(* IEC 61131-3 sources: 2026_Projet_YGO_ExcavatriceDragage/ARCHIVES/Code/PLC_TESTS/TYPES/STRUCTS, 13 files *)

(* ---- ST_PlcTestsCmd.st ---- *)
// ═══════════════════════════════════════════════════════════════
// 🧪 ST_PlcTestsCmd — Commandes de pilotage du banc de validation
// ═══════════════════════════════════════════════════════════════

TYPE ST_PlcTestsCmd :
STRUCT
    // Commandes unitaires : une seule suite manuelle à la fois.
    RunSafety     : BOOL;   // Lance la suite Safety
    RunTranslation: BOOL;   // Lance la suite Translation
    RunBucket     : BOOL;   // Lance la suite Benne
    RunEncoder    : BOOL;   // Lance la suite Codeurs/Homing
    RunModes      : BOOL;   // Lance la suite Modes/Homme-mort
    RunHeartbeat  : BOOL;   // Lance la suite Heartbeat IHM↔PLC
    RunSupervision: BOOL;   // Lance la suite Supervision/Persistance config
    RunFramework  : BOOL;   // Lance l'autotest indépendant du framework
    RunAll        : BOOL;   // Lance Safety→Translation→Bucket→Encoder→Modes→Heartbeat
    RunSuite      : INT;    // Compatibilité : >0 lance une suite manuelle
    RunCase       : INT;    // Cas de la commande unitaire sélectionnée
    Abort         : BOOL;   // Abandonne le test en cours
    ClearReport   : BOOL;   // Efface les rapports de tests
END_STRUCT
END_TYPE

(* ---- ST_PlcTestsStatus.st ---- *)
// ═══════════════════════════════════════════════════════════════
// 🧪 ST_PlcTestsStatus — États et progression des tests
// ═══════════════════════════════════════════════════════════════

TYPE ST_PlcTestsStatus :
STRUCT
    RunState         : E_TestRunState;
    SimulationActive : BOOL;       // TRUE si la simulation automate est active
    ActiveSuiteId    : INT;        // ID de la suite en cours (ex: 1)
    ActiveCaseId     : INT;        // ID du cas en cours
    ActiveStepId     : INT;        // ID de l'étape en cours
    ActiveSuiteName  : STRING(32); // Nom de la suite active
    ActiveCaseName   : STRING(32); // Nom du cas active
    ActiveStepName   : STRING(32); // Nom de l'étape active
    StepElapsed      : TIME;       // Temps écoulé dans l'étape active
    StepTimeoutPT    : TIME;       // Timeout de l'étape active
    CasesTotal       : INT;        // Nombre total de cas à jouer
    CasesPassed      : INT;        // Nombre de cas réussis
    CasesFailed      : INT;        // Nombre de cas en échec
    Heartbeat        : BOOL;       // Clignotant d'activité (3 pulses sur transition)
    FailureSummary   : STRING(255); // 🏷️ Détail des défauts du dernier run, TOUTES suites confondues (remonte Report.FailureSummary de chaque suite exécutée) — lisible sans creuser Suite*Validation
    TerminalState    : E_TestTerminalState;
    ErrorCode        : INT;
    ErrorMessage     : STRING(160);
    SuiteElapsed     : TIME;
    SuiteWatchdogExpired : BOOL;
END_STRUCT
END_TYPE

(* ---- ST_TestCaseConfig.st ---- *)
// ═══════════════════════════════════════════════════════════════
// 🧪 ST_TestCaseConfig — Configuration d'un cas de test
// ═══════════════════════════════════════════════════════════════

TYPE ST_TestCaseConfig :
STRUCT
    Name      : STRING(32);          // Libellé (ex. 'TC-01 Armement nominal')
    FirstStep : INT;                 // Première étape (SETUP) du cas de test
END_STRUCT
END_TYPE

(* ---- ST_TestCaseResult.st ---- *)
// ═══════════════════════════════════════════════════════════════
// 🧪 ST_TestCaseResult — Résultat d'un cas de test
// ═══════════════════════════════════════════════════════════════

TYPE ST_TestCaseResult :
STRUCT
    Name         : STRING(32);       // 🏷️ Libellé lisible (copié de CaseTable[i].Name) — identifie le cas sans chercher l'index
    Executed     : BOOL;             // Le cas de test a-t-elle été exécuté (ex. non exécuté si setup précédent abort)
    Ok           : BOOL;             // Succès global du cas de test
    FailedStepId : INT;              // Index de la première étape en échec (0 si aucune)
    FailReason   : E_TestFailReason; // Cause de l'échec global du cas de test
    Duration     : TIME;             // Durée totale du cas de test
END_STRUCT
END_TYPE

(* ---- ST_TestCheckConfig.st ---- *)
// ═══════════════════════════════════════════════════════════════
// 🧪 ST_TestCheckConfig — Configuration d'un check (une assertion)
// ═══════════════════════════════════════════════════════════════

TYPE ST_TestCheckConfig :
STRUCT
    Kind         : E_TestCheckKind;  // Type de check
    Mode         : E_TestCheckMode;  // Mode d'évaluation
    ProbeIdx     : INT;              // Index de la sonde dans le tableau correspondant
    ExpectedBool : BOOL;             // Valeur attendue pour BOOL_EQUAL
    ExpectedDint : DINT;             // Valeur attendue pour DINT_EQUAL / DINT_NOT_EQUAL
    ExpectedMin  : DINT;             // Bornes pour DINT_IN_RANGE
    ExpectedMax  : DINT;
    Mask         : WORD;             // Masque pour WORD_MASK_*
    RealMin      : REAL;             // Bornes pour REAL_IN_RANGE
    RealMax      : REAL;
    StablePT     : TIME;             // Durée de stabilité requise pour CHECK_WAIT_UNTIL
END_STRUCT
END_TYPE

(* ---- ST_TestEvent.st ---- *)
// 🧪 Événement journalisé par le banc de test
TYPE ST_TestEvent :
STRUCT
    Sequence       : UDINT;
    Severity       : E_TestEventSeverity;
    SuiteId        : INT;
    CaseId         : INT;
    StepId         : INT;
    Code           : INT;
    Message        : STRING(160);
END_STRUCT
END_TYPE

(* ---- ST_TestFrameworkResult.st ---- *)
// 🧪 Résultat plat de l'autotest indépendant du framework
TYPE ST_TestFrameworkResult :
STRUCT
    InProgress   : BOOL;
    AllPassed    : BOOL;
    AnyFailed    : BOOL;
    CurrentTestId: INT;
    FailedTestId : INT;
    TestsPassed  : INT;
    TestsFailed  : INT;
    ErrorMessage : STRING(160);
    RunCounter   : UDINT;
END_STRUCT
END_TYPE

(* ---- ST_TestInvariantConfig.st ---- *)
// ═══════════════════════════════════════════════════════════════
// 🧪 ST_TestInvariantConfig — Configuration d'un invariant multi-étapes
// ═══════════════════════════════════════════════════════════════

TYPE ST_TestInvariantConfig :
STRUCT
    Check          : ST_TestCheckConfig; // Configuration du check (Kind/sonde/valeur attendue)
    ArmAtStepId    : INT;                // Étape qui arme cet invariant
    DisarmAtStepId : INT;                // Étape qui désarme cet invariant (0 = jusqu'à la fin de la suite)
END_STRUCT
END_TYPE

(* ---- ST_TestStepConfig.st ---- *)
// ═══════════════════════════════════════════════════════════════
// 🧪 ST_TestStepConfig — Configuration d'une étape de test
// ═══════════════════════════════════════════════════════════════

TYPE ST_TestStepConfig :
STRUCT
    Name       : STRING(32);         // Libellé IHM + rapport
    CaseId     : INT;                // Rattachement au cas de test
    StimulusId : INT;                // Id du stimulus appliqué (0 = neutre)
    CheckIdx   : ARRAY[1..GVL_PLC_Tests_Const.MaxChecksPerStep] OF INT; // Index des checks (0 = vide)
    DwellPT    : TIME;               // Temporisation avant évaluation
    MinPT      : TIME;               // Fenêtre temporelle minimale
    TimeoutPT  : TIME;               // Temps limite pour réussir l'étape
    NextOnPass : INT;                // Étape suivante en cas de succès (0 = fin)
    NextOnFail : INT;                // Étape suivante en cas d'échec (souvent teardown, 0 = fin)
    FailAction : E_TestFailAction;   // Action en cas d'échec (continuer ou arrêter la suite)
END_STRUCT
END_TYPE

(* ---- ST_TestStepResult.st ---- *)
// ═══════════════════════════════════════════════════════════════
// 🧪 ST_TestStepResult — Résultat d'une étape de test
// ═══════════════════════════════════════════════════════════════

TYPE ST_TestStepResult :
STRUCT
    Executed          : BOOL;             // L'étape a-t-elle été exécutée ?
    Passed            : BOOL;             // L'étape a-t-elle été validée ?
    FailReason        : E_TestFailReason; // Raison de l'échec (FAIL_NONE si OK)
    FailedCheckIdx    : INT;              // Index du check fautif (0 si aucun)
    FailedInvariantId : INT;              // Index de l'invariant violé (0 si aucun)
    Duration          : TIME;             // Durée mesurée de l'étape
    ObservedBool      : BOOL;             // Valeur observée de la sonde BOOL en échec au verdict
    ObservedDint      : DINT;             // Valeur observée de la sonde DINT en échec au verdict
    ObservedReal      : REAL;             // Valeur observée de la sonde REAL en échec au verdict
END_STRUCT
END_TYPE

(* ---- ST_TestStimAnalogConfig.st ---- *)
// ═══════════════════════════════════════════════════════════════
// 🧪 ST_TestStimAnalogConfig — Configuration d'un stimulus instrumenté
// ═══════════════════════════════════════════════════════════════

TYPE ST_TestStimAnalogConfig :
STRUCT
    Kind       : E_TestStimKind;     // Type de stimulus (pulse, rampe, séquence)
    StartReal  : REAL;               // Valeur de départ pour la rampe
    TargetReal : REAL;               // Valeur cible pour la rampe
    PulsePT    : TIME;               // Durée de l'impulsion (PULSE_BOOL)
    RampPT     : TIME;               // Durée de transition de la rampe
    SeqValues  : ARRAY[1..GVL_PLC_Tests_Const.MaxSeqValues] OF REAL; // Valeurs de la séquence
    SeqCount   : INT;                // Nombre de valeurs utilisées dans la séquence
    SeqDwellPT : TIME;               // Temps de maintien de chaque valeur de la séquence
END_STRUCT
END_TYPE

(* ---- ST_TestSuiteReport.st ---- *)
// ═══════════════════════════════════════════════════════════════
// 🧪 ST_TestSuiteReport — Rapport d'une suite de tests
// ═══════════════════════════════════════════════════════════════

TYPE ST_TestSuiteReport :
STRUCT
    Name           : STRING(32);       // Nom de la suite de tests
    InProgress     : BOOL;             // Exécution en cours ?
    AllPassed      : BOOL;             // Tous les tests de la suite ont réussi ?
    AnyFailed      : BOOL;             // Au moins un échec détecté ?
    Aborted        : BOOL;             // Suite abandonnée ?
    TerminalState  : E_TestTerminalState; // 🛡️ Fin explicite, aucune attente implicite sur Done
    ErrorCode      : INT;              // Code d'erreur de configuration/exécution
    ErrorMessage   : STRING(160);      // Diagnostic court exploitable IHM/log
    FailedTestCase : INT;              // Premier cas de test en échec (0 si aucun)
    FailureSummary : STRING(255);      // 🏷️ TOUS les cas en échec en 1 ligne lisible (ex. 'TC-01 (step 15): FAIL_CHECK | TC-03 (step 30): FAIL_TIMEOUT') — évite de parcourir Cases[] un par un
    CurrentStepId  : INT;              // Étape en cours d'exécution
    CurrentCaseId  : INT;              // Cas de test en cours d'exécution
    Duration       : TIME;             // Durée totale du run de la suite
    RunCounter     : UDINT;            // Compteur de runs depuis le démarrage
    Steps          : ARRAY[1..GVL_PLC_Tests_Const.MaxSteps]     OF ST_TestStepResult;
    Cases          : ARRAY[1..GVL_PLC_Tests_Const.MaxTestCases] OF ST_TestCaseResult;
END_STRUCT
END_TYPE

(* ---- ST_TranslationTestResult.st ---- *)
// ═══════════════════════════════════════════════════════════════
// 🧪 ST_TranslationTestResult — Résultat plat de la suite Translation
// ───────────────────────────────────────────────────────────────
// 🎯 Vue synthétique lisible en 1 coup d'œil (IHM/Watch), en complément
//    du rapport détaillé existant ST_TestSuiteReport (Steps[]/Cases[]).
//    Alimenté par FB_TranslationReportFinalizer (CORE).
// ═══════════════════════════════════════════════════════════════

TYPE ST_TranslationTestResult :
STRUCT
    TerminalState    : E_TestTerminalState; // État terminal du dernier run (NONE tant qu'aucun run)
    RequestedCaseId  : INT;                 // CaseId demandé au dernier Start (0=tous, 1..6=case ciblée)
    ExecutedCaseId   : INT;                 // Dernier cas en cours/joué (0 si aucun)
    AllPassed        : BOOL;
    AnyFailed        : BOOL;
    FailedCaseId     : INT;                 // Premier cas en échec (0 = aucun)
    FailedCaseName   : STRING(32);
    FailReason       : E_TestFailReason;    // Cause du 1er cas en échec (FAIL_NONE si aucun)
    ErrorCode        : INT;
    ErrorMessage     : STRING(160);
    CasesTotal       : INT;
    CasesPassed      : INT;
    CasesFailed      : INT;
    Duration         : TIME;
    RunCounter       : UDINT;
END_STRUCT
END_TYPE
